// TIA Portal V18 export
TYPE "Udt_DataAGVStation"
   STRUCT
      Station { S7_SetPoint := 'True'} : Array[1..20] of "Udt_Data_AGVToScala";
   END_STRUCT;
END_TYPE
